FUNCTION_BLOCK TANK_HYSTERESIS (* Migrated from IEC 61131-3 ST *)
  (* Standard: 61499-2 *)
  (* Version 1.0, 2026-11-06, st2fb *)
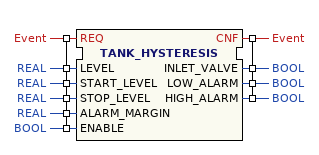
  EVENT_INPUT
    REQ WITH LEVEL, START_LEVEL, STOP_LEVEL, ALARM_MARGIN, ENABLE;
  END_EVENT
  EVENT_OUTPUT
    CNF WITH INLET_VALVE, LOW_ALARM, HIGH_ALARM;
  END_EVENT
  VAR_INPUT
    LEVEL : REAL;
    START_LEVEL : REAL;
    STOP_LEVEL : REAL;
    ALARM_MARGIN : REAL;
    ENABLE : BOOL;
  END_VAR
  VAR_OUTPUT
    INLET_VALVE : BOOL;
    LOW_ALARM : BOOL;
    HIGH_ALARM : BOOL;
  END_VAR
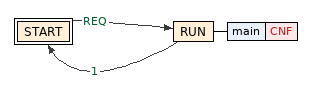
  EC_STATES
    START;
    RUN : main -> CNF;
  END_STATES
  EC_TRANSITIONS
    START TO RUN := REQ;
    RUN TO START := 1;
  END_TRANSITIONS
  ALGORITHM main IN ST:
IF NOT ENABLE THEN
  INLET_VALVE := FALSE;
ELSIF LEVEL <= START_LEVEL THEN
  INLET_VALVE := TRUE;
ELSIF LEVEL >= STOP_LEVEL THEN
  INLET_VALVE := FALSE;
END_IF;
LOW_ALARM := LEVEL < START_LEVEL - ALARM_MARGIN;
HIGH_ALARM := LEVEL > STOP_LEVEL + ALARM_MARGIN;
  END_ALGORITHM
END_FUNCTION_BLOCK
